(* Schneider Machine Expert - Basic project register_lifo_il_shared_request, file version 3.0.0.0 *)
(* ProjectInformations: Name=New project *)

HARDWARE
  Cpu 0: TM200CE40T
  EthernetConfiguration: NetworkName=M200, IpAllocationMode=FixedAddress, IpAddress=0.0.0.0, SubnetMask=0.0.0.0
  SerialLineConfiguration: Baud=Baud19200, Parity=ParityEven, DataBits=DataBits8, StopBits=StopBits1, PhysicalMedium=PhysicalMediumRs485, TransmissionMode=TransmissionModeModbusRtu, SlaveId=1, Addressing=SlaveAddressing
  MastTask: UsePeriodScanMode=false, PeriodScan=100
  FastTask: Period=255
  CpuBehavior: StartingMode=StartAsPreviousState, AutoSaveRamOnEeprom=true, WatchdogPeriod=250

SYMBOLS  (address, symbol, comment, settings)
  %R0         [Type=Lifo]

POU New POU
  (* SectionNumber=0 *)

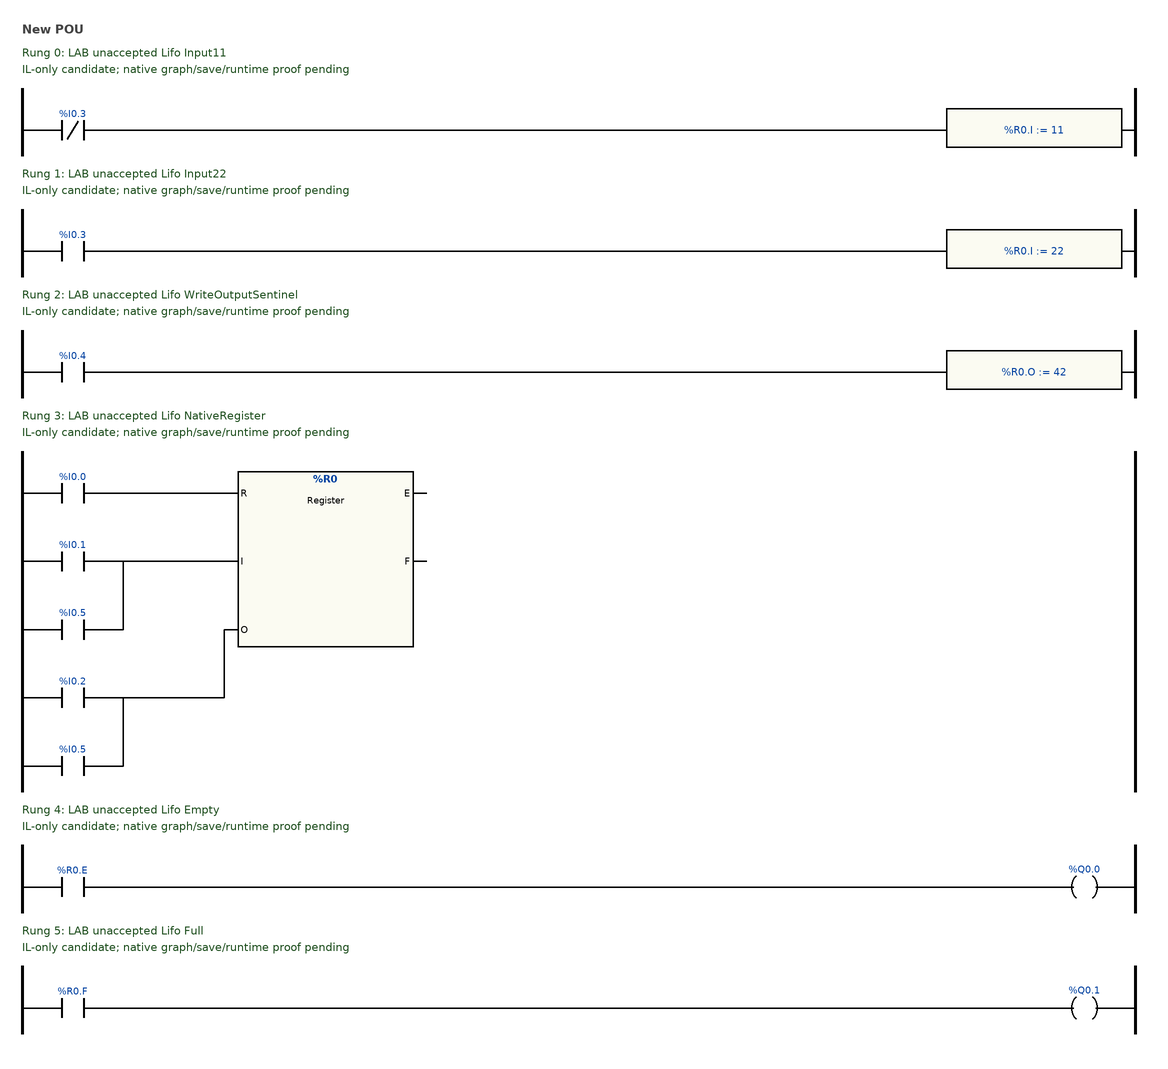

// Rung 0: LAB unaccepted Lifo Input11
// IL-only candidate; native graph/save/runtime proof pending
  LDN %I0.3
  [ %R0.I := 11 ]
  // as ST:
  //   IF NOT %I0.3 THEN %R0.I := 11; END_IF;

// Rung 1: LAB unaccepted Lifo Input22
// IL-only candidate; native graph/save/runtime proof pending
  LD %I0.3
  [ %R0.I := 22 ]
  // as ST:
  //   IF %I0.3 THEN %R0.I := 22; END_IF;

// Rung 2: LAB unaccepted Lifo WriteOutputSentinel
// IL-only candidate; native graph/save/runtime proof pending
  LD %I0.4
  [ %R0.O := 42 ]
  // as ST:
  //   IF %I0.4 THEN %R0.O := 42; END_IF;

// Rung 3: LAB unaccepted Lifo NativeRegister
// IL-only candidate; native graph/save/runtime proof pending
  BLK %R0
  LD %I0.0
  R
  LD %I0.1
  OR %I0.5
  I
  LD %I0.2
  OR %I0.5
  O
  END_BLK
  // as ST:
  //   %R0(R := %I0.0, I := %I0.1 OR %I0.5, O := %I0.2 OR %I0.5);

// Rung 4: LAB unaccepted Lifo Empty
// IL-only candidate; native graph/save/runtime proof pending
  LD %R0.E
  ST %Q0.0
  // as ST:
  //   %Q0.0 := %R0.E;

// Rung 5: LAB unaccepted Lifo Full
// IL-only candidate; native graph/save/runtime proof pending
  LD %R0.F
  ST %Q0.1
  // as ST:
  //   %Q0.1 := %R0.F;
